FUNCTION FC 1 : VOID
BEGIN
NETWORK
      A E 0.0
END_FUNCTION
